// TIA Portal V19 export
TYPE "EM05_Input"
   STRUCT
      Cmds { S7_SetPoint := 'True'} : "EM_Input";
      AgitatorType : Int := 1;   // 1=Acople superior, 2=Acople inferior
      MinLevelPermit : Bool;
   END_STRUCT;
END_TYPE
